(* IEC 61131-3 sources: trust-platform/examples/OSCAT/tunnel_washer_chain/oop/src, 3 files *)

(* ---- Main.st ---- *)
(* Record role: WasherQualityEvent is a deterministic PLC-side record for tests and runtime readers. *)
TYPE WasherQualityEvent :
STRUCT
    SoilLevel : REAL;
    Conductivity : REAL;
    RinseConductivity : REAL;
    OperatorAvailable : BOOL;
END_STRUCT
END_TYPE

(* Pattern role: IWasherQualityHandler is the contract boundary for the Chain of Responsibility example. *)
INTERFACE IWasherQualityHandler
    PROPERTY HandlerId : INT
    GET
    END_GET
    END_PROPERTY

    METHOD SetNext
    VAR_INPUT
        NextHandler : IWasherQualityHandler;
    END_VAR
    END_METHOD

    METHOD Handle : BOOL
    VAR_INPUT
        Event : WasherQualityEvent;
    END_VAR
    END_METHOD
END_INTERFACE

(* Pattern role: AutoDoseHandler is a concrete implementation in the Chain of Responsibility example. *)
FUNCTION_BLOCK AutoDoseHandler IMPLEMENTS IWasherQualityHandler
VAR
    Next : IWasherQualityHandler;
    HandledValue : BOOL;
END_VAR

METHOD PUBLIC SetNext
VAR_INPUT
    NextHandler : IWasherQualityHandler;
END_VAR
Next := NextHandler;
END_METHOD

METHOD PUBLIC Handle : BOOL
VAR_INPUT
    Event : WasherQualityEvent;
END_VAR
(* Reset on entry so HandledValue reflects only the current event. *)
HandledValue := FALSE;
IF (Event.SoilLevel > REAL#70.0) AND (Event.Conductivity < REAL#3.0) THEN
    HandledValue := TRUE;
    Handle := TRUE;
ELSE
    Handle := Next.Handle(Event := Event);
END_IF;
END_METHOD

PUBLIC PROPERTY HandlerId : INT
GET
    HandlerId := INT#1;
END_GET
END_PROPERTY

PUBLIC PROPERTY Handled : BOOL
GET
    Handled := HandledValue;
END_GET
END_PROPERTY
END_FUNCTION_BLOCK

(* Pattern role: ExtendRinseHandler is a concrete implementation in the Chain of Responsibility example. *)
FUNCTION_BLOCK ExtendRinseHandler IMPLEMENTS IWasherQualityHandler
VAR
    Next : IWasherQualityHandler;
    HandledValue : BOOL;
END_VAR

METHOD PUBLIC SetNext
VAR_INPUT
    NextHandler : IWasherQualityHandler;
END_VAR
Next := NextHandler;
END_METHOD

METHOD PUBLIC Handle : BOOL
VAR_INPUT
    Event : WasherQualityEvent;
END_VAR
(* Reset on entry so HandledValue reflects only the current event. *)
HandledValue := FALSE;
IF Event.RinseConductivity > REAL#1.5 THEN
    HandledValue := TRUE;
    Handle := TRUE;
ELSE
    Handle := Next.Handle(Event := Event);
END_IF;
END_METHOD

PUBLIC PROPERTY HandlerId : INT
GET
    HandlerId := INT#2;
END_GET
END_PROPERTY

PUBLIC PROPERTY Handled : BOOL
GET
    Handled := HandledValue;
END_GET
END_PROPERTY
END_FUNCTION_BLOCK

(* Pattern role: OperatorHoldHandler is a concrete implementation in the Chain of Responsibility example. *)
FUNCTION_BLOCK OperatorHoldHandler IMPLEMENTS IWasherQualityHandler
VAR
    Next : IWasherQualityHandler;
    HandledValue : BOOL;
END_VAR

METHOD PUBLIC SetNext
VAR_INPUT
    NextHandler : IWasherQualityHandler;
END_VAR
Next := NextHandler;
END_METHOD

METHOD PUBLIC Handle : BOOL
VAR_INPUT
    Event : WasherQualityEvent;
END_VAR
(* Reset on entry so HandledValue reflects only the current event. *)
HandledValue := FALSE;
IF Event.OperatorAvailable THEN
    HandledValue := TRUE;
    Handle := TRUE;
ELSE
    Handle := Next.Handle(Event := Event);
END_IF;
END_METHOD

PUBLIC PROPERTY HandlerId : INT
GET
    HandlerId := INT#3;
END_GET
END_PROPERTY

PUBLIC PROPERTY Handled : BOOL
GET
    Handled := HandledValue;
END_GET
END_PROPERTY
END_FUNCTION_BLOCK

(* Pattern role: RejectBatchHandler is a concrete implementation in the Chain of Responsibility example. *)
FUNCTION_BLOCK RejectBatchHandler IMPLEMENTS IWasherQualityHandler
VAR
    HandledValue : BOOL;
END_VAR

METHOD PUBLIC SetNext
VAR_INPUT
    NextHandler : IWasherQualityHandler;
END_VAR
END_METHOD

METHOD PUBLIC Handle : BOOL
VAR_INPUT
    Event : WasherQualityEvent;
END_VAR
(* Last handler in the chain: always handles. Reset on entry so the
   flag reflects only this event. *)
HandledValue := TRUE;
Handle := TRUE;
END_METHOD

PUBLIC PROPERTY HandlerId : INT
GET
    HandlerId := INT#4;
END_GET
END_PROPERTY

PUBLIC PROPERTY Handled : BOOL
GET
    Handled := HandledValue;
END_GET
END_PROPERTY
END_FUNCTION_BLOCK

(* Composition role: TunnelWasherQualityController owns the collaborating objects used by this Chain of Responsibility example. *)
FUNCTION_BLOCK TunnelWasherQualityController
VAR
    AutoDose : AutoDoseHandler;
    ExtendRinse : ExtendRinseHandler;
    OperatorHold : OperatorHoldHandler;
    RejectBatch : RejectBatchHandler;
    Chain : IWasherQualityHandler;
    AutoDoseCounter : DwordCounter;
    RejectCounter : DwordCounter;
    LastHandlerIdValue : INT;
END_VAR

METHOD PUBLIC Initialize
AutoDose.SetNext(NextHandler := ExtendRinse);
ExtendRinse.SetNext(NextHandler := OperatorHold);
OperatorHold.SetNext(NextHandler := RejectBatch);
Chain := AutoDose;
AutoDoseCounter.Initialize();
AutoDoseCounter.Configure(StepSize := DWORD#1, MaxValue := DWORD#16#FFFFFFFF);
RejectCounter.Initialize();
RejectCounter.Configure(StepSize := DWORD#1, MaxValue := DWORD#16#FFFFFFFF);
END_METHOD

METHOD PUBLIC Evaluate : INT
VAR_INPUT
    SoilLevel : REAL;
    Conductivity : REAL;
    RinseConductivity : REAL;
    OperatorAvailable : BOOL;
END_VAR
VAR
    Event : WasherQualityEvent;
END_VAR
Event.SoilLevel := SoilLevel;
Event.Conductivity := Conductivity;
Event.RinseConductivity := RinseConductivity;
Event.OperatorAvailable := OperatorAvailable;
(* DwordCounter wraps COUNT_DR which is edge-triggered (UP AND NOT
   LastUp). Drop the UP edge first so consecutive same-class events
   each generate a fresh rising edge and actually increment. *)
AutoDoseCounter.Update(Up := FALSE, Down := FALSE);
RejectCounter.Update(Up := FALSE, Down := FALSE);
Chain.Handle(Event := Event);
IF AutoDose.Handled THEN
    LastHandlerIdValue := AutoDose.HandlerId;
    AutoDoseCounter.Update(Up := TRUE, Down := FALSE);
ELSIF ExtendRinse.Handled THEN
    LastHandlerIdValue := ExtendRinse.HandlerId;
ELSIF OperatorHold.Handled THEN
    LastHandlerIdValue := OperatorHold.HandlerId;
ELSE
    LastHandlerIdValue := RejectBatch.HandlerId;
    RejectCounter.Update(Up := TRUE, Down := FALSE);
END_IF;
Evaluate := LastHandlerIdValue;
END_METHOD

PUBLIC PROPERTY LastHandlerId : INT
GET
    LastHandlerId := LastHandlerIdValue;
END_GET
END_PROPERTY

PUBLIC PROPERTY RejectCount : DWORD
GET
    RejectCount := RejectCounter.Count;
END_GET
END_PROPERTY

PUBLIC PROPERTY AutoDoseCount : DWORD
GET
    AutoDoseCount := AutoDoseCounter.Count;
END_GET
END_PROPERTY
END_FUNCTION_BLOCK

(* Scan role: Main wires the example objects and exposes the PLC call path under test. *)
PROGRAM Main
VAR
    Washer : TunnelWasherQualityController;
    SoilLevelRaw : INT;
    ConductivityRaw : INT;
    OperatorAvailable : BOOL;
    DosePumpOut : BOOL;
    RejectOut : BOOL;
END_VAR

Washer.Initialize();
Washer.Evaluate(SoilLevel := INT_TO_REAL(SoilLevelRaw), Conductivity := INT_TO_REAL(ConductivityRaw) / REAL#10.0, RinseConductivity := REAL#0.8, OperatorAvailable := OperatorAvailable);
DosePumpOut := Washer.LastHandlerId = INT#1;
RejectOut := Washer.LastHandlerId = INT#4;
END_PROGRAM

(* ---- Configuration.st ---- *)
CONFIGURATION TunnelWasherChainOopConfiguration
RESOURCE TunnelWasherChainOop ON PLC
    TASK MainTask (INTERVAL := T#100ms, PRIORITY := 1);
    PROGRAM Washer WITH MainTask : Main;
END_RESOURCE
VAR_CONFIG
    Washer.SoilLevelRaw AT %IW2 : INT;
    Washer.ConductivityRaw AT %IW4 : INT;
    Washer.OperatorAvailable AT %IX0.0 : BOOL;
    Washer.DosePumpOut AT %QX0.0 : BOOL;
    Washer.RejectOut AT %QX0.1 : BOOL;
END_VAR
END_CONFIGURATION

(* ---- Tests.st ---- *)
TEST_PROGRAM WasherChainStopsAtAutoDose
VAR
    Washer : TunnelWasherQualityController;
END_VAR

Washer.Initialize();
ASSERT_EQUAL(EXPECTED := INT#1, ACTUAL := Washer.Evaluate(SoilLevel := REAL#80.0, Conductivity := REAL#2.0, RinseConductivity := REAL#0.5, OperatorAvailable := FALSE));
ASSERT_EQUAL(EXPECTED := DWORD#1, ACTUAL := Washer.AutoDoseCount);
END_TEST_PROGRAM

TEST_PROGRAM WasherChainFallsThroughToReject
VAR
    Washer : TunnelWasherQualityController;
END_VAR

Washer.Initialize();
ASSERT_EQUAL(EXPECTED := INT#4, ACTUAL := Washer.Evaluate(SoilLevel := REAL#40.0, Conductivity := REAL#4.0, RinseConductivity := REAL#0.5, OperatorAvailable := FALSE));
ASSERT_EQUAL(EXPECTED := DWORD#1, ACTUAL := Washer.RejectCount);
END_TEST_PROGRAM

(* Stale-flag regression test: drives multiple events through one
   Washer instance with different paths. Catches the bug where a
   handler keeps reporting "I handled it" after the first event
   because HandledValue is not reset on entry to Handle. *)
TEST_PROGRAM WasherChainHandlerFlagsResetBetweenEvaluations
VAR
    Washer : TunnelWasherQualityController;
END_VAR

Washer.Initialize();

(* Event 1: AutoDose path - high soil, low conductivity *)
ASSERT_EQUAL(EXPECTED := INT#1, ACTUAL := Washer.Evaluate(SoilLevel := REAL#80.0, Conductivity := REAL#2.0, RinseConductivity := REAL#0.5, OperatorAvailable := FALSE));

(* Event 2: must fall through to RejectBatch. Without the per-call
   reset of HandledValue, this returns INT#1 because AutoDose.Handled
   is still TRUE from Event 1. *)
ASSERT_EQUAL(EXPECTED := INT#4, ACTUAL := Washer.Evaluate(SoilLevel := REAL#40.0, Conductivity := REAL#4.0, RinseConductivity := REAL#0.5, OperatorAvailable := FALSE));

(* Event 3: ExtendRinse path *)
ASSERT_EQUAL(EXPECTED := INT#2, ACTUAL := Washer.Evaluate(SoilLevel := REAL#40.0, Conductivity := REAL#4.0, RinseConductivity := REAL#2.0, OperatorAvailable := FALSE));

(* Event 4: must fall through to Reject again *)
ASSERT_EQUAL(EXPECTED := INT#4, ACTUAL := Washer.Evaluate(SoilLevel := REAL#40.0, Conductivity := REAL#4.0, RinseConductivity := REAL#0.5, OperatorAvailable := FALSE));

(* Counters: 1 auto-dose, 2 rejects across the four events *)
ASSERT_EQUAL(EXPECTED := DWORD#1, ACTUAL := Washer.AutoDoseCount);
ASSERT_EQUAL(EXPECTED := DWORD#2, ACTUAL := Washer.RejectCount);
END_TEST_PROGRAM

(* AutoDoseHandler in isolation: tests the AND of two conditions. *)
TEST_PROGRAM AutoDoseHandlerHandlesOnlyHighSoilLowConductivity
VAR
    Handler : AutoDoseHandler;
    Terminal : RejectBatchHandler;
    Event : WasherQualityEvent;
END_VAR
Handler.SetNext(NextHandler := Terminal);

(* Both conditions met: handles *)
Event.SoilLevel := REAL#80.0;
Event.Conductivity := REAL#2.0;
Event.RinseConductivity := REAL#0.5;
Event.OperatorAvailable := FALSE;
Handler.Handle(Event := Event);
ASSERT_TRUE(IN := Handler.Handled);

(* Soil too low: passes through *)
Event.SoilLevel := REAL#50.0;
Handler.Handle(Event := Event);
ASSERT_FALSE(IN := Handler.Handled);

(* Conductivity too high: passes through *)
Event.SoilLevel := REAL#80.0;
Event.Conductivity := REAL#5.0;
Handler.Handle(Event := Event);
ASSERT_FALSE(IN := Handler.Handled);

(* Boundary: soil exactly 70 - strict greater-than required *)
Event.SoilLevel := REAL#70.0;
Event.Conductivity := REAL#2.0;
Handler.Handle(Event := Event);
ASSERT_FALSE(IN := Handler.Handled);

(* Boundary: conductivity exactly 3 - strict less-than required *)
Event.SoilLevel := REAL#80.0;
Event.Conductivity := REAL#3.0;
Handler.Handle(Event := Event);
ASSERT_FALSE(IN := Handler.Handled);
END_TEST_PROGRAM

(* ExtendRinseHandler: triggers on RinseConductivity > 1.5. *)
TEST_PROGRAM ExtendRinseHandlerHandlesAboveRinseThreshold
VAR
    Handler : ExtendRinseHandler;
    Terminal : RejectBatchHandler;
    Event : WasherQualityEvent;
END_VAR
Handler.SetNext(NextHandler := Terminal);

(* Above threshold: handles *)
Event.RinseConductivity := REAL#2.0;
Handler.Handle(Event := Event);
ASSERT_TRUE(IN := Handler.Handled);

(* At threshold (strict greater-than): passes through *)
Event.RinseConductivity := REAL#1.5;
Handler.Handle(Event := Event);
ASSERT_FALSE(IN := Handler.Handled);

(* Below threshold: passes through *)
Event.RinseConductivity := REAL#0.5;
Handler.Handle(Event := Event);
ASSERT_FALSE(IN := Handler.Handled);
END_TEST_PROGRAM

(* OperatorHoldHandler: triggers when OperatorAvailable. *)
TEST_PROGRAM OperatorHoldHandlerHandlesWhenOperatorAvailable
VAR
    Handler : OperatorHoldHandler;
    Terminal : RejectBatchHandler;
    Event : WasherQualityEvent;
END_VAR
Handler.SetNext(NextHandler := Terminal);

Event.OperatorAvailable := TRUE;
Handler.Handle(Event := Event);
ASSERT_TRUE(IN := Handler.Handled);

Event.OperatorAvailable := FALSE;
Handler.Handle(Event := Event);
ASSERT_FALSE(IN := Handler.Handled);
END_TEST_PROGRAM

(* RejectBatchHandler: always handles regardless of event. *)
TEST_PROGRAM RejectBatchHandlerAlwaysHandles
VAR
    Handler : RejectBatchHandler;
    Event : WasherQualityEvent;
END_VAR
Event.SoilLevel := REAL#0.0;
Event.Conductivity := REAL#0.0;
Event.RinseConductivity := REAL#0.0;
Event.OperatorAvailable := FALSE;
ASSERT_TRUE(IN := Handler.Handle(Event := Event));
ASSERT_TRUE(IN := Handler.Handled);

(* Even with all conditions favoring upstream handlers, terminal still handles *)
Event.SoilLevel := REAL#100.0;
Event.Conductivity := REAL#1.0;
Event.RinseConductivity := REAL#5.0;
Event.OperatorAvailable := TRUE;
ASSERT_TRUE(IN := Handler.Handle(Event := Event));
END_TEST_PROGRAM

(* Counter accumulation across many events. *)
TEST_PROGRAM WasherCountersAccumulateCorrectlyAcrossManyEvents
VAR
    Washer : TunnelWasherQualityController;
END_VAR
Washer.Initialize();

(* 3 auto-dose events *)
Washer.Evaluate(SoilLevel := REAL#80.0, Conductivity := REAL#2.0, RinseConductivity := REAL#0.5, OperatorAvailable := FALSE);
Washer.Evaluate(SoilLevel := REAL#85.0, Conductivity := REAL#1.0, RinseConductivity := REAL#0.5, OperatorAvailable := FALSE);
Washer.Evaluate(SoilLevel := REAL#90.0, Conductivity := REAL#0.5, RinseConductivity := REAL#0.5, OperatorAvailable := FALSE);
ASSERT_EQUAL(EXPECTED := DWORD#3, ACTUAL := Washer.AutoDoseCount);

(* 2 reject events *)
Washer.Evaluate(SoilLevel := REAL#40.0, Conductivity := REAL#5.0, RinseConductivity := REAL#0.5, OperatorAvailable := FALSE);
Washer.Evaluate(SoilLevel := REAL#30.0, Conductivity := REAL#5.0, RinseConductivity := REAL#0.5, OperatorAvailable := FALSE);
ASSERT_EQUAL(EXPECTED := DWORD#3, ACTUAL := Washer.AutoDoseCount);
ASSERT_EQUAL(EXPECTED := DWORD#2, ACTUAL := Washer.RejectCount);

(* ExtendRinse and OperatorHold do not increment AutoDose or Reject *)
Washer.Evaluate(SoilLevel := REAL#40.0, Conductivity := REAL#5.0, RinseConductivity := REAL#2.0, OperatorAvailable := FALSE);
Washer.Evaluate(SoilLevel := REAL#40.0, Conductivity := REAL#5.0, RinseConductivity := REAL#0.5, OperatorAvailable := TRUE);
ASSERT_EQUAL(EXPECTED := DWORD#3, ACTUAL := Washer.AutoDoseCount);
ASSERT_EQUAL(EXPECTED := DWORD#2, ACTUAL := Washer.RejectCount);
END_TEST_PROGRAM
